// TIA Portal V20 export
TYPE "T_DISCON_DATA"
   STRUCT
      TDISCON : Struct
         IN : Struct
            DISCONNECT : Bool;
            ID : CONN_OUC;
         END_STRUCT;
         OUT : Struct
            DONE : Bool;
            BUSY : Bool;
            ERROR : Bool;
            STATUS : Word;
         END_STRUCT;
      END_STRUCT;
   END_STRUCT;
END_TYPE
